TYPE ST_Slot :
STRUCT
    bOccupied : BOOL;
    sLeId     : STRING(20);   // load unit id (pallet barcode)
    bTaught   : BOOL;         // TRUE once the place was measured in teach mode
    lrTaughtX : LREAL;        // measured travel position [m]
    lrTaughtY : LREAL;        // measured hoist position [m]
END_STRUCT
END_TYPE

(* stored: Version 1.1.0.1
   DUT ST_Slot: Id {49e7efe3-08fb-4b4d-9ecf-adbb9a774f2a} *)
